Yaskawa INFORM job: TAKEPAR.JBI

/JOB
//NAME TAKEPAR
//POS
///NPOS 3,0,0,0,0,0
///TOOL 9
///POSTYPE PULSE
///PULSE
C00000=-74,-4,-62,162,-60,-81
///TOOL 9
///POSTYPE BASE
///RECTAN
///RCONF 1,0,0,0,0,0,0,0
C00001=290.000,-1755.000,230.000,90.00,-0.00,0.00
///RCONF 0,0,0,0,0,0,0,0
C00002=290.000,-1755.000,810.000,90.00,-0.00,0.00
//INST
///DATE 2026/10/26 01:19
///COMM Generated using RoboDK
///ATTR SC,RW,RJ
///GROUP1 RB1
NOP
'Using Table (targets wrt base
'):
'0.0,-1500.0,-60.0,0.0,0.0,0.0
'Setting Tool 9 (Wood_Holder):
SETE P00095 (1) 0
SETE P00095 (2) 0
SETE P00095 (3) 40000
SETE P00095 (4) 0
SETE P00095 (5) 0
SETE P00095 (6) 0
SETTOOL TL#(9) P00095
MOVJ C00000 VJ=50.00
MOVL C00001 V=1000.0
'Attach to Wood_Holder
'Attach to Wood_Holder
MOVL C00002 V=1000.0
END
